(* Test host that nests an FB_SLITS_POWER, the way a device FB would. Its references and
   values are bound in its own FB_Init, which runs after the nested FB_SLITS_POWER was
   constructed from them, so the nested FB_SLITS_POWER first sees nil references and
   empty values. CallAfterInit re-supplies all of them through
   fbSlits.CallAfterInitPOWER. *)
{attribute 'call_after_init'}
FUNCTION_BLOCK FB_SLITSPOWERHost
VAR
    {attribute 'no_copy'}
    aiMotionStage : REFERENCE TO ARRAY[1..4] OF I_MotionStage;
    {attribute 'no_copy'}
    fbFFHWO       : REFERENCE TO FB_HardwareFFOutput;
    sDeviceName   : STRING;
    bBridgeOK     : REFERENCE TO BOOL;
    sPmpsState    : STRING;
    {attribute 'no_copy'}
    bFileReaderBusy : REFERENCE TO BOOL;
    fApertureMargin : REAL;
    bBridgeConfirmedBad : REFERENCE TO BOOL;

    fbSlits : FB_SLITS_POWER(
        aiMotionStage   := aiMotionStage,
        fbFFHWO         := fbFFHWO,
        sDeviceName     := sDeviceName,
        bBridgeOK       := bBridgeOK,
        sPmpsState      := sPmpsState,
        bFileReaderBusy := bFileReaderBusy,
        fApertureMargin := fApertureMargin,
        bBridgeConfirmedBad := bBridgeConfirmedBad
    );
END_VAR

fbSlits(
    bMoveOk := TRUE
);

(* The nested fbSlits ran its own CallAfterInit before this one, with nil
   references. Re-supplies them and redoes its wiring. *)
{attribute 'call_after_init'}
METHOD CallAfterInit
fbSlits.CallAfterInitPOWER(
    aiMotionStage   := aiMotionStage,
    fbFFHWO         := fbFFHWO,
    sDeviceName     := sDeviceName,
    bBridgeOK       := bBridgeOK,
    sPmpsState      := sPmpsState,
    bFileReaderBusy := bFileReaderBusy,
    fApertureMargin := fApertureMargin,
    bBridgeConfirmedBad := bBridgeConfirmedBad
);
END_METHOD

(* Stores the injected references and values in this FB's fields. *)
{attribute 'analysis' := '-33'}
METHOD FB_Init : BOOL
VAR_INPUT
    bInitRetains : BOOL;
    bInCopyCode  : BOOL;
    aiMotionStage : REFERENCE TO ARRAY[1..4] OF I_MotionStage;
    fbFFHWO       : REFERENCE TO FB_HardwareFFOutput;
    sDeviceName   : STRING;
    bBridgeOK     : REFERENCE TO BOOL;
    sPmpsState    : STRING;
    bFileReaderBusy : REFERENCE TO BOOL;
    fApertureMargin : REAL;
    bBridgeConfirmedBad : REFERENCE TO BOOL;
END_VAR
THIS^.aiMotionStage REF= aiMotionStage;
THIS^.fbFFHWO       REF= fbFFHWO;
THIS^.sDeviceName   := sDeviceName;
THIS^.bBridgeOK     REF= bBridgeOK;
THIS^.sPmpsState    := sPmpsState;
THIS^.bFileReaderBusy REF= bFileReaderBusy;
THIS^.fApertureMargin := fApertureMargin;
THIS^.bBridgeConfirmedBad REF= bBridgeConfirmedBad;
END_METHOD

(* Sets the per-blade encoder zero-offsets of the nested slit, which are inputs
   of the slit that only this host can reach. *)
METHOD SetEncoderOffsets
VAR_INPUT
    Top    : REAL;
    Bottom : REAL;
    North  : REAL;
    South  : REAL;
END_VAR
fbSlits.rEncoderOffsetTop    := Top;
fbSlits.rEncoderOffsetBottom := Bottom;
fbSlits.rEncoderOffsetNorth  := North;
fbSlits.rEncoderOffsetSouth  := South;
END_METHOD

(* Requests a gap and a centre from the nested slit, as an EPICS write would. *)
METHOD SetAperture
VAR_INPUT
    SizeX   : REAL;
    SizeY   : REAL;
    CenterX : REAL;
    CenterY : REAL;
END_VAR
fbSlits.SetApertureRequest(
    ApertureSizeX := SizeX,
    ApertureSizeY := SizeY,
    CenterX       := CenterX,
    CenterY       := CenterY
);
END_METHOD

(* Stands in for the PMPS aperture the arbiter would send: sets the request that
   becomes the trusted limit, so a larger gap request is accepted. *)
METHOD SetTrustedAperture
VAR_INPUT
    Width  : REAL;
    Height : REAL;
END_VAR
fbSlits.SetAptWidthHeight(
    Width  := Width,
    Height := Height
);
END_METHOD

(* Runs the PMPS aperture reconciliation of the nested power slit, as a power-slit
   program does each cycle. Index is the slit's slot in astApertures. *)
METHOD UpdatePMPS
VAR_INPUT
    Index : INT;
END_VAR
fbSlits.M_UpdatePMPS(
    index := Index
);
END_METHOD

END_FUNCTION_BLOCK

(* stored: Version 1.1.0.1
   POU FB_SLITSPOWERHost: Id {8c1b91a6-ca7f-4a02-bc9c-34a7fd009c26}, SpecialFunc None
   Method CallAfterInit: Id {775acb7f-9335-40e0-87d6-c4b0615fc8dc}
   Method FB_Init: Id {d5efdb8b-7ef0-46ca-b164-f00bbe6ac779}
   Method SetEncoderOffsets: Id {a56e5279-5ec1-4a86-b991-4ef261d76613}
   Method SetAperture: Id {e80bceeb-44da-43d5-a5fe-318e76c10592}
   Method SetTrustedAperture: Id {cd585572-2ee4-43ac-908b-f7be0ffbdff3}
   Method UpdatePMPS: Id {fc8088b8-38f2-4646-9a55-60052e6f7a17} *)
